Fanuc KAREL source: KD00066.KL

PROGRAM KD00066
%NOLOCKGROUP
VAR
  I: INTEGER
  J: INTEGER
  B: BOOLEAN
  R: REAL
  S: STRING[80]
BEGIN
  CONDITION[1]:
  WHEN DIN[1] = ON DO
    NOPAUSE
  ENDCONDITION
END KD00066
